(* PMPS-aware (power-class) variant of FB_SLITS. Adds 8 thermocouple RTDs,
   a flow switch, a reactive-temp DB lookup (FB_JsonDocToSafeBP keyed by
   sPmpsState) driving every RTD fault, an xPMPSMode toggle, and M_UpdatePMPS.
   EXTENDS FB_SLITS; body calls SUPER^() for edge-trigger consumption then
   drives M_CalculatePositions / M_Motion behind a REF nil-guard. *)
{attribute 'analysis' := '-33'}
{attribute 'call_after_init'}
FUNCTION_BLOCK FB_SLITS_POWER EXTENDS FB_SLITS

VAR
    {attribute 'pytmc' := '
    pv: MODE
    field: ZNAM Local
    field: ONAM PMPS
    io: io
    '}
    xPMPSMode : BOOL := TRUE;

    {attribute 'pytmc' := 'pv: FSW'}
    fbFlowSwitch : FB_XTES_Flowswitch;

    {attribute 'pytmc' := 'pv: TOP:RTD:01'}
    RTD_TOP_1 : FB_CC_TempSensor;
    {attribute 'pytmc' := 'pv: TOP:RTD:02'}
    RTD_TOP_2 : FB_CC_TempSensor;
    {attribute 'pytmc' := 'pv: BOTTOM:RTD:01'}
    RTD_Bottom_1 : FB_CC_TempSensor;
    {attribute 'pytmc' := 'pv: BOTTOM:RTD:02'}
    RTD_Bottom_2 : FB_CC_TempSensor;
    {attribute 'pytmc' := 'pv: NORTH:RTD:01'}
    RTD_North_1 : FB_CC_TempSensor;
    {attribute 'pytmc' := 'pv: NORTH:RTD:02'}
    RTD_North_2 : FB_CC_TempSensor;
    {attribute 'pytmc' := 'pv: SOUTH:RTD:01'}
    RTD_South_1 : FB_CC_TempSensor;
    {attribute 'pytmc' := 'pv: SOUTH:RTD:02'}
    RTD_South_2 : FB_CC_TempSensor;
    (* PMPS reactive-DB key for the device's allowed temperature. *)
    sPmpsState : STRING;
    fbReadPMPSDB : FB_JsonDocToSafeBP;
    astTempDB    : ARRAY[1..1] OF ST_DbStateParams;
    (* fbReadPMPSDB.bExecute needs a rising edge; a real PMPS file read produces one as bBusy falls.
       Taken as REFERENCE TO so a test can drive its own BOOL and simulate the edge
       instead of reaching into MOTION_GVL.fbPmpsFileReader directly.
    *)
    bFileReaderBusy : REFERENCE TO BOOL;
    (* Margin (mm) subtracted from the authorized width/height when snapping
       the request into PMPS compliance. Set via FB_Init, defaults to 0.01. *)
    fApertureMargin : REAL := 0.01;
END_VAR

IF NOT __ISVALIDREF(THIS^.aiMotionStage)
   OR NOT __ISVALIDREF(THIS^.fbFFHWO) OR NOT __ISVALIDREF(bFileReaderBusy) THEN
    RETURN;
END_IF


// Parent body: EPICS edge-trigger consumption only (no REF touch).
SUPER^();


// Inherited dispatch (parity with legacy FB_SLITS_POWER body
// invoking ACT_CalculatePositions / ACT_Motion).
M_CalculatePositions();
M_Motion();

// PMPS reactive temperature DB lookup. bExecute needs a rising edge,
// produced as the caller-injected file-reader busy flag falls. Guard
// the REF (single condition, no short-circuit hazard) so an unbound
// instance stays inert rather than dereferencing a nil ref.
astTempDB[1].sPmpsState := sPmpsState;
fbReadPMPSDB(
    bExecute    := NOT bFileReaderBusy,
    jsonDoc     := PMPS_GVL.BP_jsonDoc,
    sDeviceName := sDeviceName,
    arrStates   := astTempDB,
    io_fbFFHWO  := fbFFHWO
);

// All 8 RTDs share the same fault threshold (resolved from the DB).
RTD_TOP_1(
    fFaultThreshold := astTempDB[1].stReactiveParams.nTempSP,
    sDevName        := sDeviceName,
    io_fbFFHWO      := fbFFHWO
);
RTD_TOP_2(
    fFaultThreshold := astTempDB[1].stReactiveParams.nTempSP,
    sDevName        := sDeviceName,
    io_fbFFHWO      := fbFFHWO
);
RTD_Bottom_1(
    fFaultThreshold := astTempDB[1].stReactiveParams.nTempSP,
    sDevName        := sDeviceName,
    io_fbFFHWO      := fbFFHWO
);
RTD_Bottom_2(
    fFaultThreshold := astTempDB[1].stReactiveParams.nTempSP,
    sDevName        := sDeviceName,
    io_fbFFHWO      := fbFFHWO
);
RTD_North_1(
    fFaultThreshold := astTempDB[1].stReactiveParams.nTempSP,
    sDevName        := sDeviceName,
    io_fbFFHWO      := fbFFHWO
);
RTD_North_2(
    fFaultThreshold := astTempDB[1].stReactiveParams.nTempSP,
    sDevName        := sDeviceName,
    io_fbFFHWO      := fbFFHWO
);
RTD_South_1(
    fFaultThreshold := astTempDB[1].stReactiveParams.nTempSP,
    sDevName        := sDeviceName,
    io_fbFFHWO      := fbFFHWO
);
RTD_South_2(
    fFaultThreshold := astTempDB[1].stReactiveParams.nTempSP,
    sDevName        := sDeviceName,
    io_fbFFHWO      := fbFFHWO
);

fbFlowSwitch();

(* Records sPmpsState and REF-binds the caller-owned file-reader busy flag;
   aiMotionStage (4 blades), fbFFHWO and sDeviceName are bound by base
   FB_SLITS.FB_Init. Blade wiring runs from CallAfterInit. *)
{attribute 'analysis' := '-33'}
METHOD FB_Init : BOOL
VAR_INPUT
    bInitRetains  : BOOL;
    bInCopyCode   : BOOL;
    aiMotionStage : REFERENCE TO ARRAY[1..4] OF I_MotionStage;
    fbFFHWO       : REFERENCE TO FB_HardwareFFOutput;
    sDeviceName   : STRING;
    sPmpsState 	  : STRING;
    bFileReaderBusy : REFERENCE TO BOOL;
    fApertureMargin : REAL;
END_VAR
THIS^.sPmpsState := sPmpsState;
THIS^.bFileReaderBusy REF= bFileReaderBusy;
THIS^.fApertureMargin := fApertureMargin;
END_METHOD

(* Integrator-driven PMPS aperture-safety reconciliation, called each cycle
   with index = this device's slot in astApertures. Mirrors actual geometry
   into AptArrayStatus, faults FFO when actual gap exceeds the authorized
   envelope (or always, out of PMPS mode), and in PMPS mode snaps the request
   into compliance. Caller must ensure index is valid (no short-circuit). *)
METHOD M_UpdatePMPS : BOOL
VAR_INPUT
    index : INT;
END_VAR
// Mirror current actual aperture geometry and any-blade error state.
THIS^.AptArrayStatus.Height := THIS^.rActApertureSizeY;
THIS^.AptArrayStatus.Width  := THIS^.rActApertureSizeX;
THIS^.AptArrayStatus.xOK    :=
        NOT (THIS^.aiMotionStage[E_SlitsBlade.TOP   ].MotionStatus.bError)
    AND NOT (THIS^.aiMotionStage[E_SlitsBlade.BOTTOM].MotionStatus.bError)
    AND NOT (THIS^.aiMotionStage[E_SlitsBlade.NORTH ].MotionStatus.bError)
    AND NOT (THIS^.aiMotionStage[E_SlitsBlade.SOUTH ].MotionStatus.bError);

// Aperture-envelope evaluation.
IF ( THIS^.rActApertureSizeX > (AptArrayReq.Width  - (2 * ABS(THIS^.rActCenterX)))
     AND PMPS_GVL.stCurrentBeamParameters.astApertures[index].Width  > 0 )
OR ( THIS^.rActApertureSizeY > (AptArrayReq.Height - (2 * ABS(THIS^.rActCenterY)))
     AND PMPS_GVL.stCurrentBeamParameters.astApertures[index].Height > 0 ) THEN
    FFO.i_xOK := FALSE;
ELSE
    FFO.i_xOK := TRUE;
END_IF

IF xPMPSMode THEN
    IF THIS^.rActApertureSizeX > AptArrayReq.Width THEN
        rReqApertureSizeX := AptArrayReq.Width - fApertureMargin;
    END_IF
    IF THIS^.rActApertureSizeY > AptArrayReq.Height THEN
        rReqApertureSizeY := AptArrayReq.Height - fApertureMargin;
    END_IF
ELSE
    FFO.i_xOK := FALSE;
END_IF

FFO(
    i_xAutoReset := TRUE,
    io_fbFFHWO   := fbFFHWO
);
END_METHOD

END_FUNCTION_BLOCK

(* stored: Version 1.1.0.1
   POU FB_SLITS_POWER: Id {f2a7b61c-c24f-40b8-8c2e-4d94fdfd3c86}, SpecialFunc None
   Method FB_Init: Id {374dff7e-a7f7-48ec-a96e-6c5ba3e1db5a}
   Method M_UpdatePMPS: Id {d82078ab-8935-40b4-85a2-97a1fdb15da8} *)
